(* IEC 61131-3 sources: plcassist-cli/packages/volt-lsp-iec/test-corpus/pro2193/Device/Plc Logic/Application/99 Library/Functions/PositionReached, 2 files *)

(* ---- PositionReached.fun ---- *)
// Check if two positions match (within 1 mm).
FUNCTION PositionReached : BOOL
VAR_INPUT
	rActPos		: REAL;
	rSetPos		: REAL;
END_VAR

PositionReached			:= PositionReachedValue(rActPos, rSetPos, 1);

END_FUNCTION

(* ---- PositionReachedValue.fun ---- *)
// Check if two positions match (within rValue mm).
FUNCTION PositionReachedValue : BOOL
VAR_INPUT
	rActPos		: REAL;
	rSetPos		: REAL;
	rValue		: REAL;
END_VAR

PositionReachedValue	:= ABS(rActPos - rSetPos) <= rValue;

END_FUNCTION
